Staubli VAL3: bind.pgx

program bind()
  local string l_sbtn
  local num l_i
begin
  //button
  userPageBindClick("editProg","btnback",bBack,true)
  for l_i = 1 to 8
    l_sbtn="btn"+toString("",l_i)
    userPageBindClick("editProg",l_sbtn,bBool[l_i],true)
  endFor

  for l_i = 0 to 8
    l_sbtn="btn1"+toString("",l_i)
    userPageBindClick("editProg",l_sbtn,bInsert[l_i],true)
  endFor

  //lbl
  userPageBind("editProg","lbl1","innerHTML",sSelProg,1,"r")
  userPageBind("editProg","lbleditindex","innerHTML",sPageIndex,1,"r")
  userPageBind("editProg","lbleditpage","innerHTML",sPageNum,1,"r")

  //lst
  userPageBind("editProg","lst1","options",sList,size(sList),"r")
  userPageBind("editProg","lst1","value",sLstValue,1,"rw")

end
